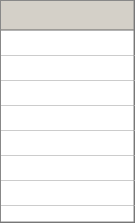
VISUALIZATION Vis_PauseHistory  // 135x223
VAR_IN_OUT
	fbOp: FB_Operation;
END_VAR
    Table (0,0 135x223), data array: fbOp.arPauseHistory
        p3854506369: fbOp.arPauseHistory[INDEX]
        p2232123230: Pause History
END_VISUALIZATION

(* stored: Version 1.1.0.1, ProductVersion 3.1.4024.13
   Visu Vis_PauseHistory: Id {c77094e4-90f3-4f67-bcf3-7187fabe8132} *)
